TEXTLIST TextList_Piston_Recipe_State_OnOff
  0 = ' '
  1 = 'On'
  2 = 'Off'
   = ''
END_TEXTLIST

(* stored: Version 1.1.0.1, ProductVersion 3.1.4024.12
   TextList TextList_Piston_Recipe_State_OnOff: Id {b6dd1aa4-2b34-4e98-9385-ae04369e151b} *)
